// TIA Portal V21 export
VAR_GLOBAL   // PLC tag table "Sensorik"
   di_axis_ref_h AT %I2.7 : Bool;
   di_axis_ref_v AT %I2.6 : Bool;
END_VAR
